// CFC twin of T_SafeRTrig_UserFB_Tests: the same tests drawn as CFC diagrams, the way a TwinSAFE project is authored.
    FUNCTION_BLOCK T_SafeRTrig_UserFB_Tests_CFC EXTENDS T_SafeCfcTestSuite
    VAR
    // Test_TriggerForOneCycleOnRisingEdge
    group_1 : T_SafeGroup;
    fb_1 : T_SafeRTrig_UserFB(group := group_1);
    // Test_StoppedGivesNoOutput
    group_2 : T_SafeGroup;
    fb_2 : T_SafeRTrig_UserFB(group := group_2);
    // Test_InnerBlocksJoinTheGroup
    group_3 : T_SafeGroup;
    fb_3 : T_SafeRTrig_UserFB(group := group_3);
END_VAR

Test_TriggerForOneCycleOnRisingEdge();
Test_StoppedGivesNoOutput();
Test_InnerBlocksJoinTheGroup();

METHOD PRIVATE Test_InnerBlocksJoinTheGroup
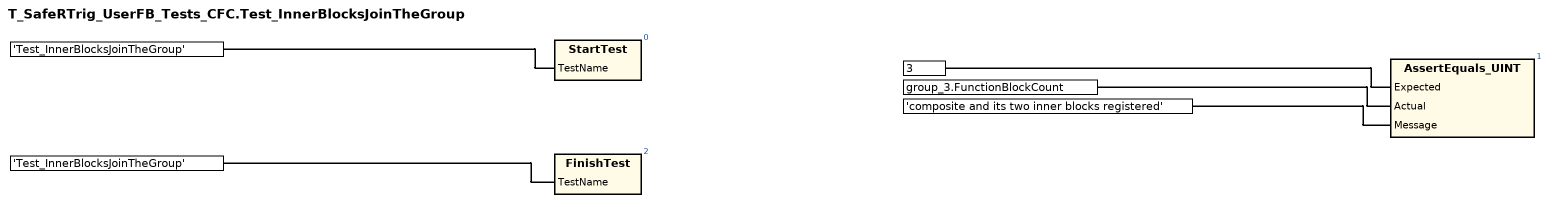
StartTest(TestName := 'Test_InnerBlocksJoinTheGroup');
AssertEquals_UINT(Expected := 3, Actual := group_3.FunctionBlockCount, Message := 'composite and its two inner blocks registered');
FinishTest(TestName := 'Test_InnerBlocksJoinTheGroup');
END_METHOD

METHOD PRIVATE Test_StoppedGivesNoOutput
// note: this text did not pass the execution check against the stored diagram
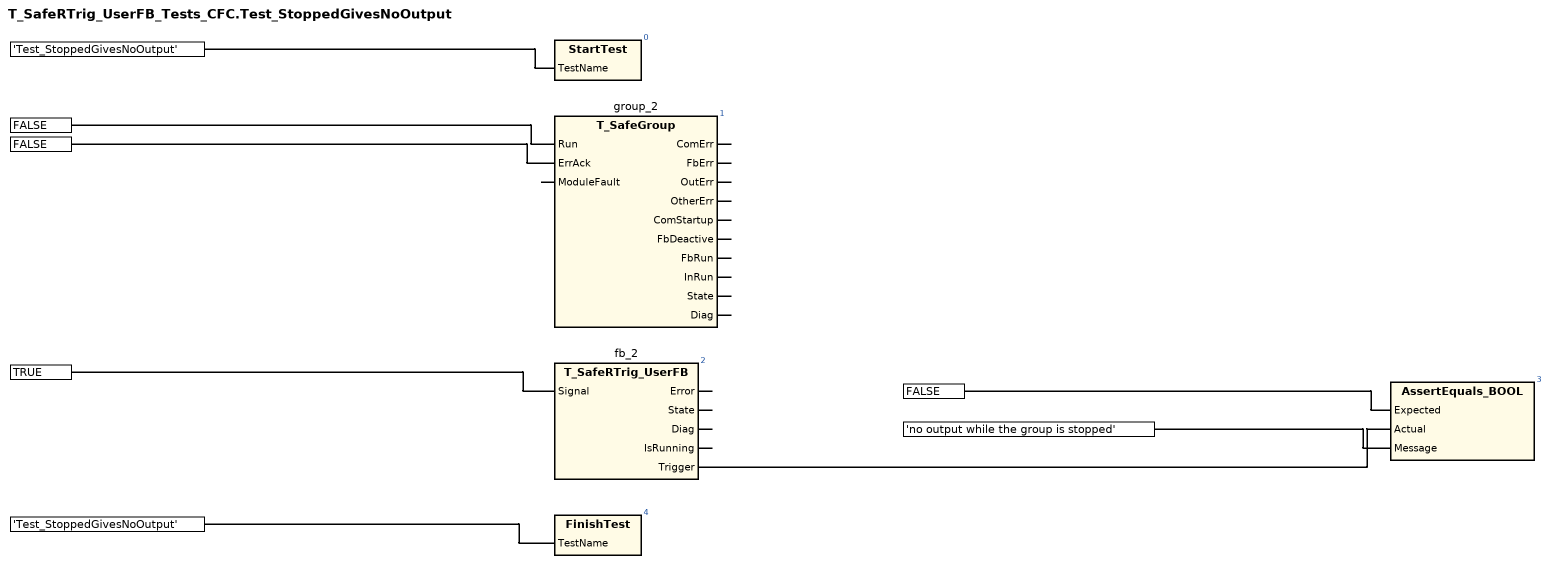
StartTest(TestName := 'Test_StoppedGivesNoOutput');
group_2(Run := FALSE, ErrAck := FALSE); // T_SafeGroup
fb_2(Signal := TRUE); // T_SafeRTrig_UserFB
AssertEquals_BOOL(Expected := FALSE, Actual := fb_2.Trigger, Message := 'no output while the group is stopped');
FinishTest(TestName := 'Test_StoppedGivesNoOutput');
END_METHOD

METHOD PRIVATE Test_TriggerForOneCycleOnRisingEdge
// note: this text did not pass the execution check against the stored diagram
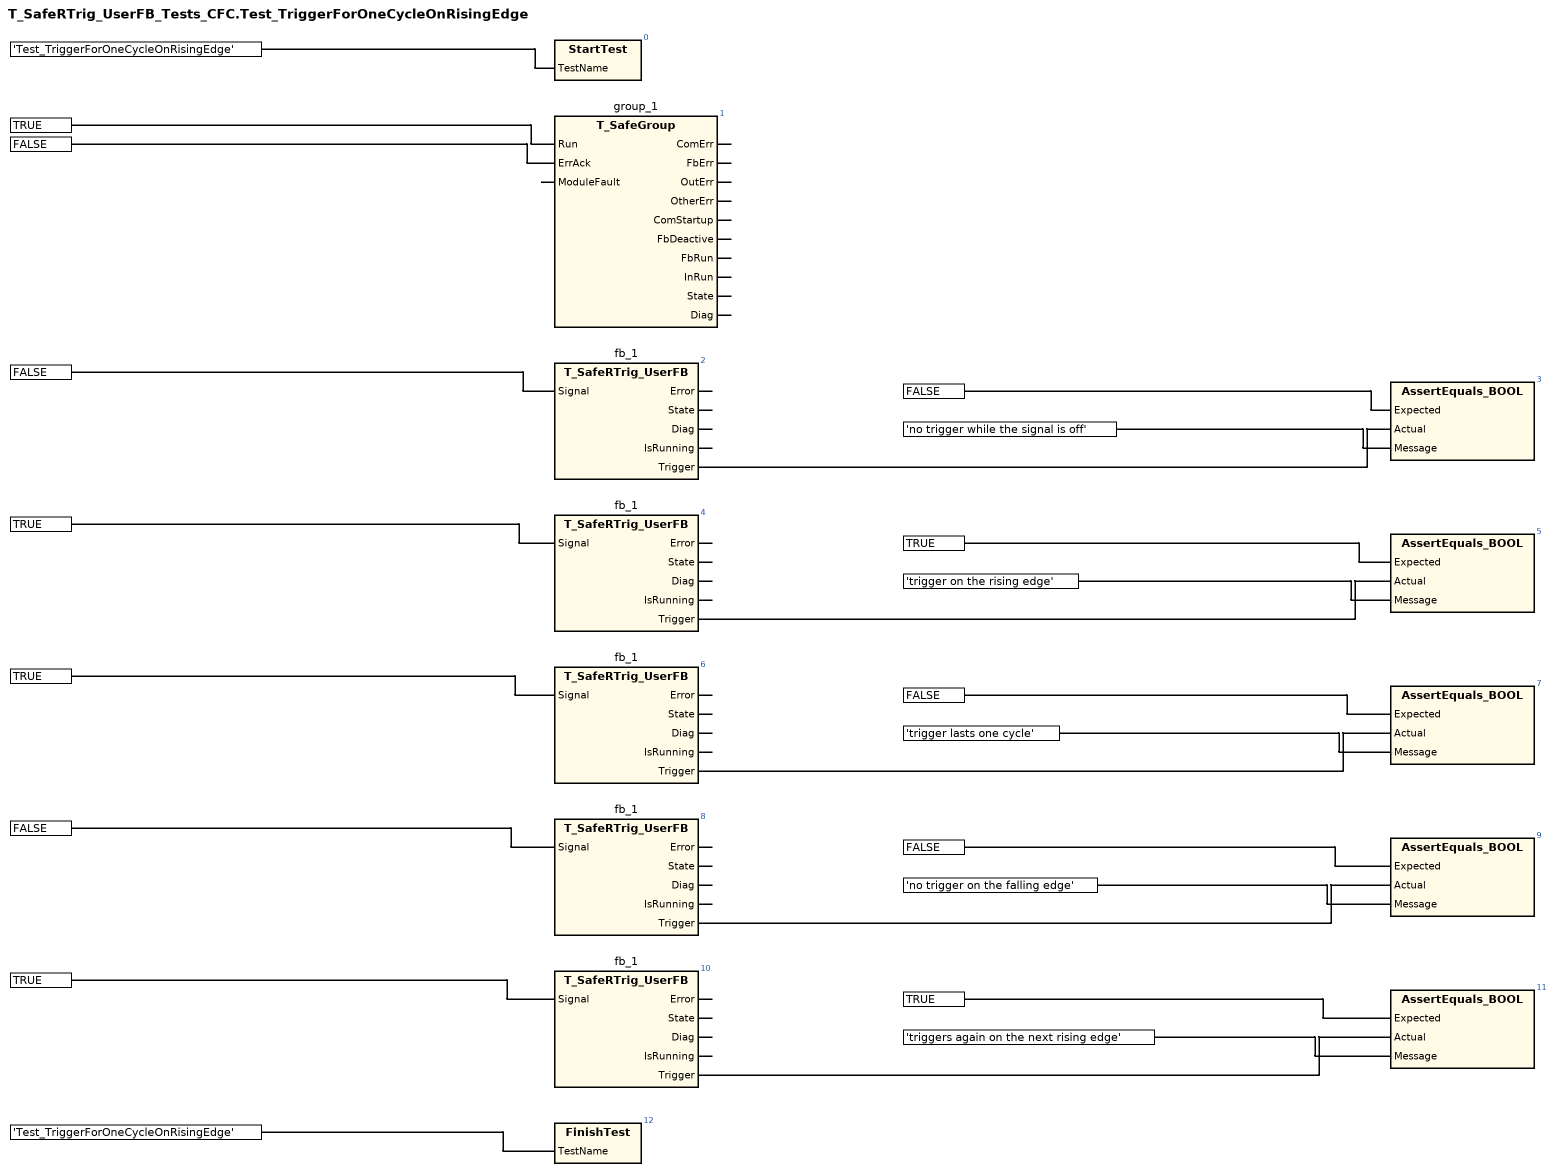
StartTest(TestName := 'Test_TriggerForOneCycleOnRisingEdge');
group_1(Run := TRUE, ErrAck := FALSE); // T_SafeGroup
fb_1(Signal := FALSE); // T_SafeRTrig_UserFB
AssertEquals_BOOL(Expected := FALSE, Actual := fb_1.Trigger, Message := 'no trigger while the signal is off');
fb_1(Signal := TRUE); // T_SafeRTrig_UserFB
AssertEquals_BOOL(Expected := TRUE, Actual := fb_1.Trigger, Message := 'trigger on the rising edge');
fb_1(Signal := TRUE); // T_SafeRTrig_UserFB
AssertEquals_BOOL(Expected := FALSE, Actual := fb_1.Trigger, Message := 'trigger lasts one cycle');
fb_1(Signal := FALSE); // T_SafeRTrig_UserFB
AssertEquals_BOOL(Expected := FALSE, Actual := fb_1.Trigger, Message := 'no trigger on the falling edge');
fb_1(Signal := TRUE); // T_SafeRTrig_UserFB
AssertEquals_BOOL(Expected := TRUE, Actual := fb_1.Trigger, Message := 'triggers again on the next rising edge');
FinishTest(TestName := 'Test_TriggerForOneCycleOnRisingEdge');
END_METHOD

END_FUNCTION_BLOCK

(* stored: Version 1.1.0.1
   POU T_SafeRTrig_UserFB_Tests_CFC: Id {6bab9a86-ad8c-5de3-9a5a-59b7d0175202}, SpecialFunc None
   Method Test_InnerBlocksJoinTheGroup: Id {fe627fee-ff97-5185-99e7-02b3fcf52b36}
   Method Test_StoppedGivesNoOutput: Id {c13ec495-5bff-5c50-8253-12f172da57cd}
   Method Test_TriggerForOneCycleOnRisingEdge: Id {963ecec9-b5f4-5218-891c-3947889ea87a} *)
